FUNCTION F_CycleSec : REAL		// 지금 태스크의 주기 (s)
VAR
	nTask		: DINT;
END_VAR

nTask := GETCURTASKINDEXEX();
F_CycleSec := UDINT_TO_REAL(TwinCAT_SystemInfoVarList._TaskInfo[nTask].CycleTime) * 1.0E-7;	// 100 ns 단위

END_FUNCTION

(* stored: Version 1.1.0.1, ProductVersion 3.1.4024.15
   POU F_CycleSec: Id {8a7384bc-b606-4438-bdf5-f5576645071c}, SpecialFunc None *)
